(* PLC project g_comb_or, Anonymous Benchmark Suite 1.0 *)
(* stored: creationDateTime 2026-08-26T00:00:00 *)

PROGRAM g_comb_or
  VAR_INPUT
    A : BOOL;
    B : BOOL;
  END_VAR
  VAR_OUTPUT
    Y : BOOL;
  END_VAR

(* LD diagram, written out as Structured Text *)
Y := A OR B;
END_PROGRAM

CONFIGURATION Config0
  RESOURCE Res0 ON PLC
    TASK tcyclic(INTERVAL := T#10ms, PRIORITY := 0);
    PROGRAM inst0 WITH tcyclic : g_comb_or;
  END_RESOURCE
END_CONFIGURATION
